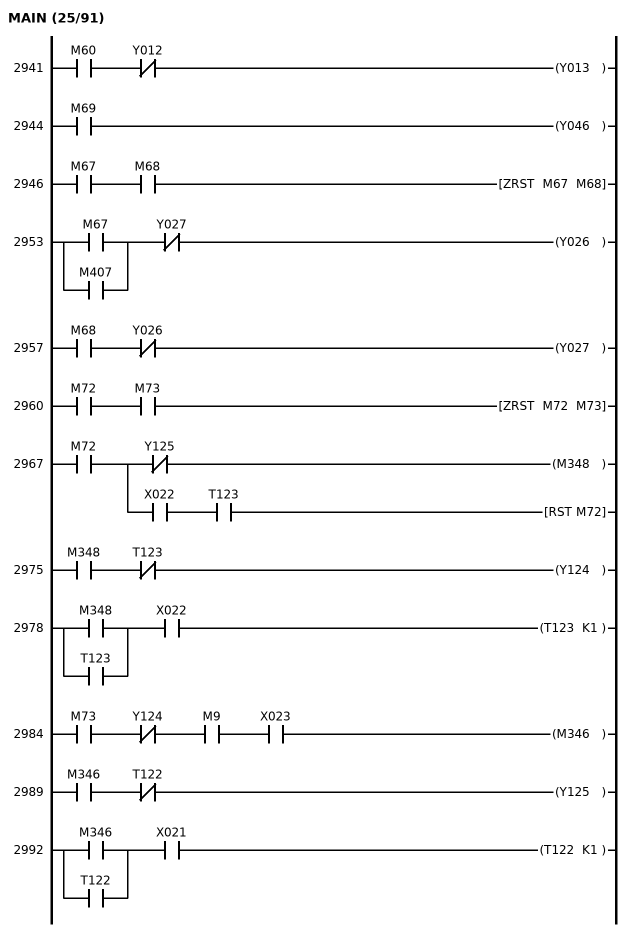
[picture p24: ladder of MAIN, rungs at steps 2941 to 2992]
2941  LD      M60
      ANI     Y012
      OUT     Y013
2944  LD      M69
      OUT     Y046
2946  LD      M67
      AND     M68
      ZRST    M67 M68
2953  LD      M67
      OR      M407
      ANI     Y027
      OUT     Y026
2957  LD      M68
      ANI     Y026
      OUT     Y027
2960  LD      M72
      AND     M73
      ZRST    M72 M73
2967  LD      M72
      MPS
      ANI     Y125
      OUT     M348
      MPP
      AND     X022
      AND     T123
      RST     M72
2975  LD      M348
      ANI     T123
      OUT     Y124
2978  LD      M348
      OR      T123
      AND     X022
      OUT     T123 K1
2984  LD      M73
      ANI     Y124
      AND     M9
      AND     X023
      OUT     M346
2989  LD      M346
      ANI     T122
      OUT     Y125
2992  LD      M346
      OR      T122
      AND     X021
      OUT     T122 K1
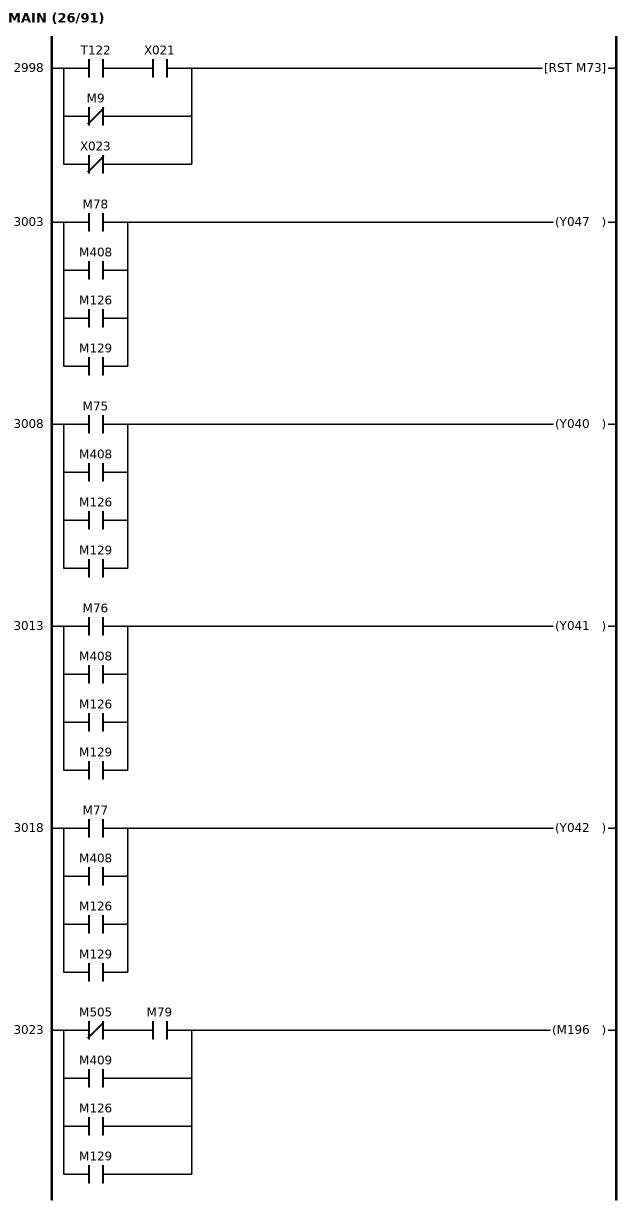
2998  LD      T122
      AND     X021
      ORI     M9
      ORI     X023
      RST     M73
3003  LD      M78
      OR      M408
      OR      M126
      OR      M129
      OUT     Y047
3008  LD      M75
      OR      M408
      OR      M126
      OR      M129
      OUT     Y040
3013  LD      M76
      OR      M408
      OR      M126
      OR      M129
      OUT     Y041
3018  LD      M77
      OR      M408
      OR      M126
      OR      M129
      OUT     Y042
3023  LDI     M505
      AND     M79
      OR      M409
      OR      M126
      OR      M129
      OUT     M196
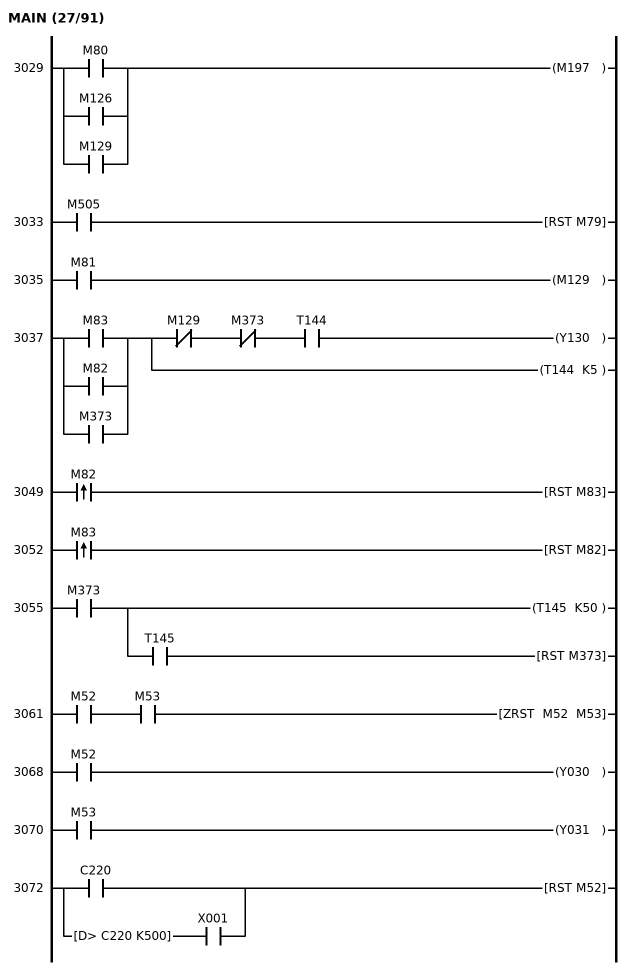
3029  LD      M80
      OR      M126
      OR      M129
      OUT     M197
3033  LD      M505
      RST     M79
3035  LD      M81
      OUT     M129
3037  LD      M83
      OR      M82
      OR      M373
      MPS
      ANI     M129
      ANI     M373
      AND     T144
      OUT     Y130
      MPP
      OUT     T144 K5
3049  LDP     M82
      RST     M83
3052  LDP     M83
      RST     M82
3055  LD      M373
      OUT     T145 K50
      AND     T145
      RST     M373
3061  LD      M52
      AND     M53
      ZRST    M52 M53
3068  LD      M52
      OUT     Y030
3070  LD      M53
      OUT     Y031
3072  LD      C220
      LDD>    C220 K500
      AND     X001
      ORB
      RST     M52
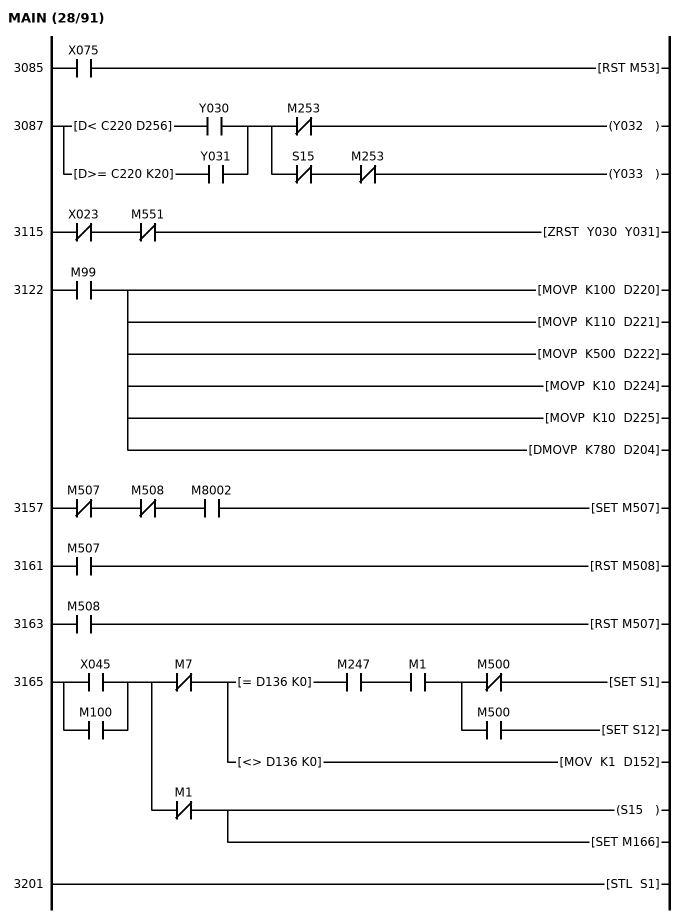
3085  LD      X075
      RST     M53
3087  LDD<    C220 D256
      AND     Y030
      LDD>=   C220 K20
      AND     Y031
      ORB
      MPS
      ANI     M253
      OUT     Y032
      MPP
      ANI     S15
      ANI     M253
      OUT     Y033
3115  LDI     X023
      ANI     M551
      ZRST    Y030 Y031
3122  LD      M99
      MOVP    K100 D220
      MOVP    K110 D221
      MOVP    K500 D222
      MOVP    K10 D224
      MOVP    K10 D225
      DMOVP   K780 D204
3157  LDI     M507
      ANI     M508
      AND     M8002
      SET     M507
3161  LD      M507
      RST     M508
3163  LD      M508
      RST     M507
3165  LD      X045
      OR      M100
      MPS
      ANI     M7
      MPS
      AND=    D136 K0
      AND     M247
      AND     M1
      MPS
      ANI     M500
      SET     S1
      MPP
      AND     M500
      SET     S12
      MPP
      AND<>   D136 K0
      MOV     K1 D152
      MPP
      ANI     M1
      OUT     S15
      SET     M166
3201  STL     S1
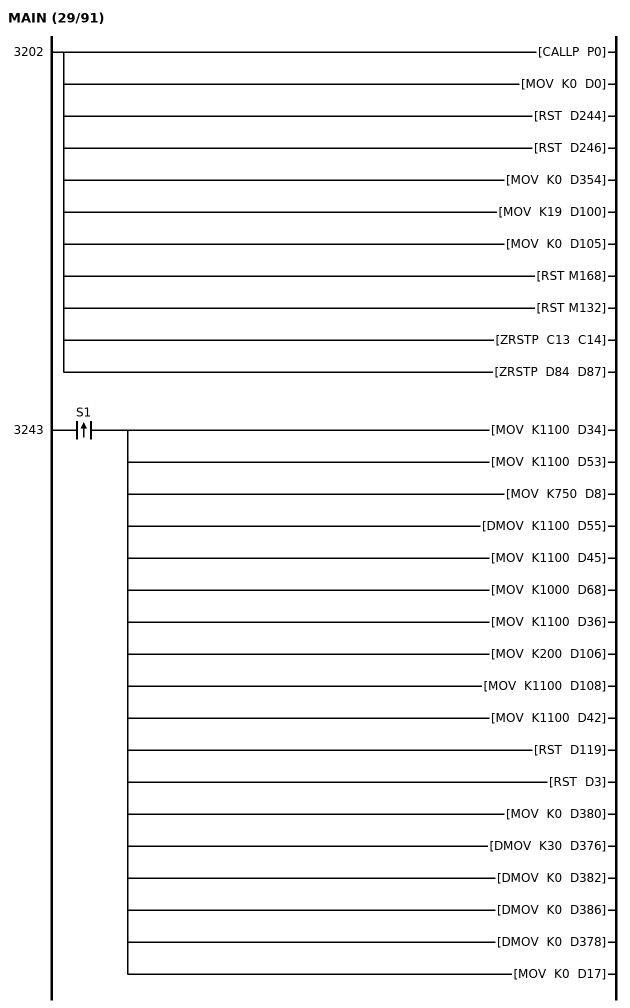
3202  CALLP   P0
      MOV     K0 D0
      RST     D244
      RST     D246
      MOV     K0 D354
      MOV     K19 D100
      MOV     K0 D105
      RST     M168
      RST     M132
      ZRSTP   C13 C14
      ZRSTP   D84 D87
3243  LDP     S1
      MOV     K1100 D34
      MOV     K1100 D53
      MOV     K750 D8
      DMOV    K1100 D55
      MOV     K1100 D45
      MOV     K1000 D68
      MOV     K1100 D36
      MOV     K200 D106
      MOV     K1100 D108
      MOV     K1100 D42
      RST     D119
      RST     D3
      MOV     K0 D380
      DMOV    K30 D376
      DMOV    K0 D382
      DMOV    K0 D386
      DMOV    K0 D378
      MOV     K0 D17
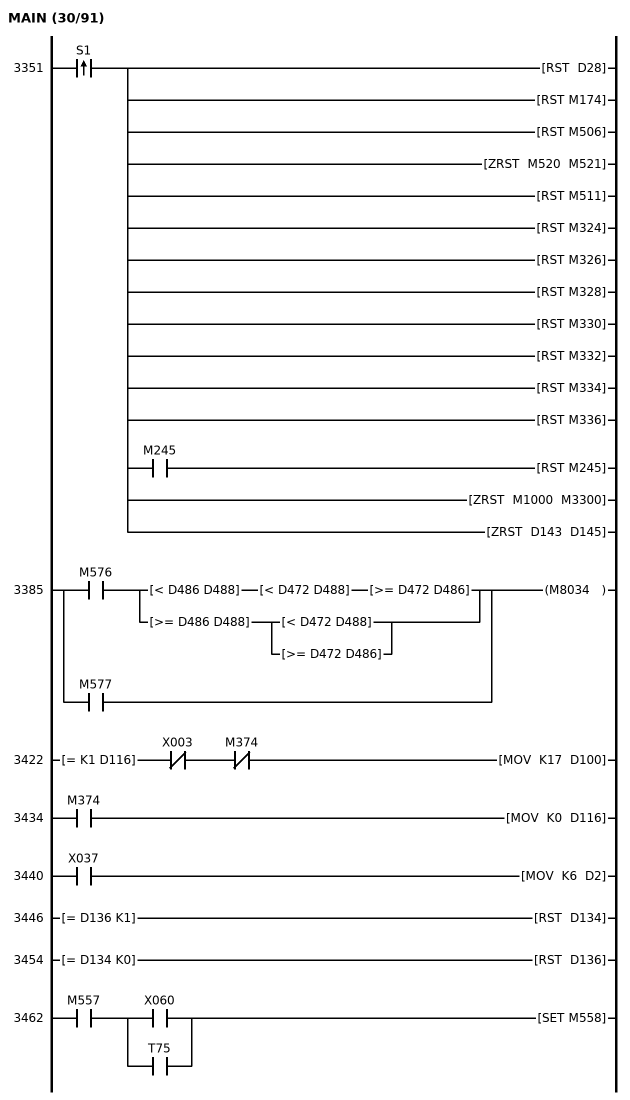
3351  LDP     S1
      RST     D28
      RST     M174
      RST     M506
      ZRST    M520 M521
      RST     M511
      RST     M324
      RST     M326
      RST     M328
      RST     M330
      RST     M332
      RST     M334
      RST     M336
      MPS
      AND     M245
      RST     M245
      MPP
      ZRST    M1000 M3300
      ZRST    D143 D145
3385  LD      M576
      LD<     D486 D488
      AND<    D472 D488
      AND>=   D472 D486
      LD>=    D486 D488
      LD<     D472 D488
      OR>=    D472 D486
      ANB
      ORB
      ANB
      OR      M577
      OUT     M8034
3422  LD=     K1 D116
      ANI     X003
      ANI     M374
      MOV     K17 D100
3434  LD      M374
      MOV     K0 D116
3440  LD      X037
      MOV     K6 D2
3446  LD=     D136 K1
      RST     D134
3454  LD=     D134 K0
      RST     D136
3462  LD      M557
      LD      X060
      OR      T75
      ANB
      SET     M558
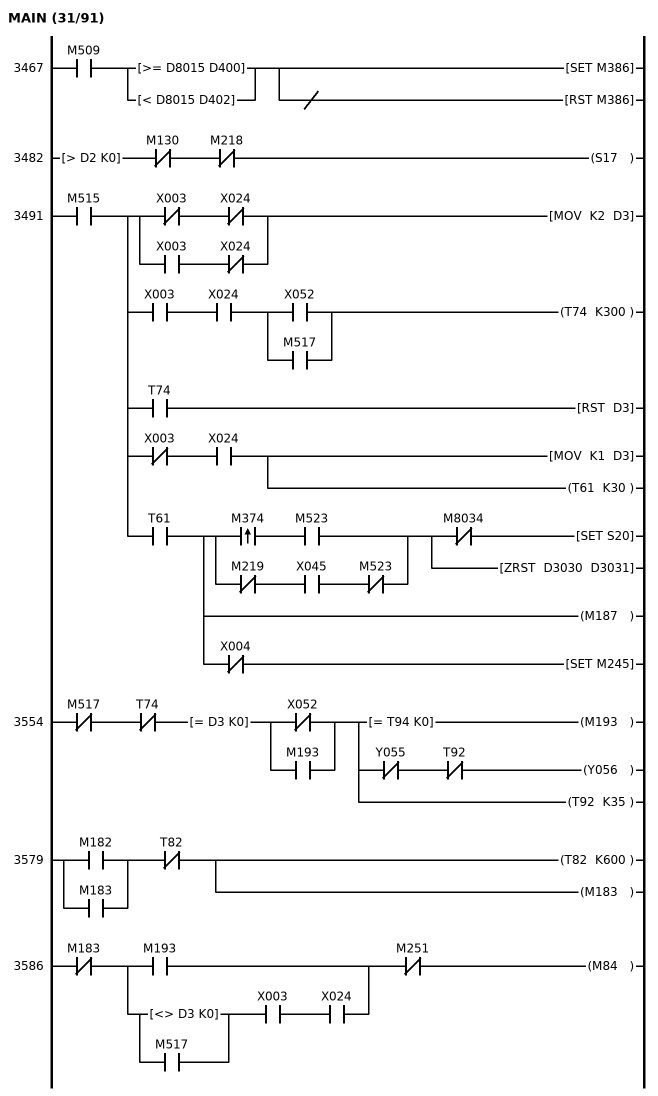
3467  LD      M509
      LD>=    D8015 D400
      OR<     D8015 D402
      ANB
      SET     M386
      INV
      RST     M386
3482  LD>     D2 K0
      ANI     M130
      ANI     M218
      OUT     S17
3491  LD      M515
      MPS
      LDI     X003
      ANI     X024
      LD      X003
      ANI     X024
      ORB
      ANB
      MOV     K2 D3
      MRD
      AND     X003
      AND     X024
      LD      X052
      OR      M517
      ANB
      OUT     T74 K300
      MRD
      AND     T74
      RST     D3
      MRD
      ANI     X003
      AND     X024
      MOV     K1 D3
      OUT     T61 K30
      MPP
      AND     T61
      MPS
      LDP     M374
      AND     M523
      LDI     M219
      AND     X045
      ANI     M523
      ORB
      ANB
      MPS
      ANI     M8034
      SET     S20
      MPP
      ZRST    D3030 D3031
      MPP
      OUT     M187
      ANI     X004
      SET     M245
3554  LDI     M517
      ANI     T74
      AND=    D3 K0
      LDI     X052
      OR      M193
      ANB
      MPS
      AND=    T94 K0
      OUT     M193
      MRD
      ANI     Y055
      ANI     T92
      OUT     Y056
      MPP
      OUT     T92 K35
3579  LD      M182
      OR      M183
      ANI     T82
      OUT     T82 K600
      OUT     M183
3586  LDI     M183
      LD      M193
      LD<>    D3 K0
      OR      M517
      AND     X003
      AND     X024
      ORB
      ANB
      ANI     M251
      OUT     M84
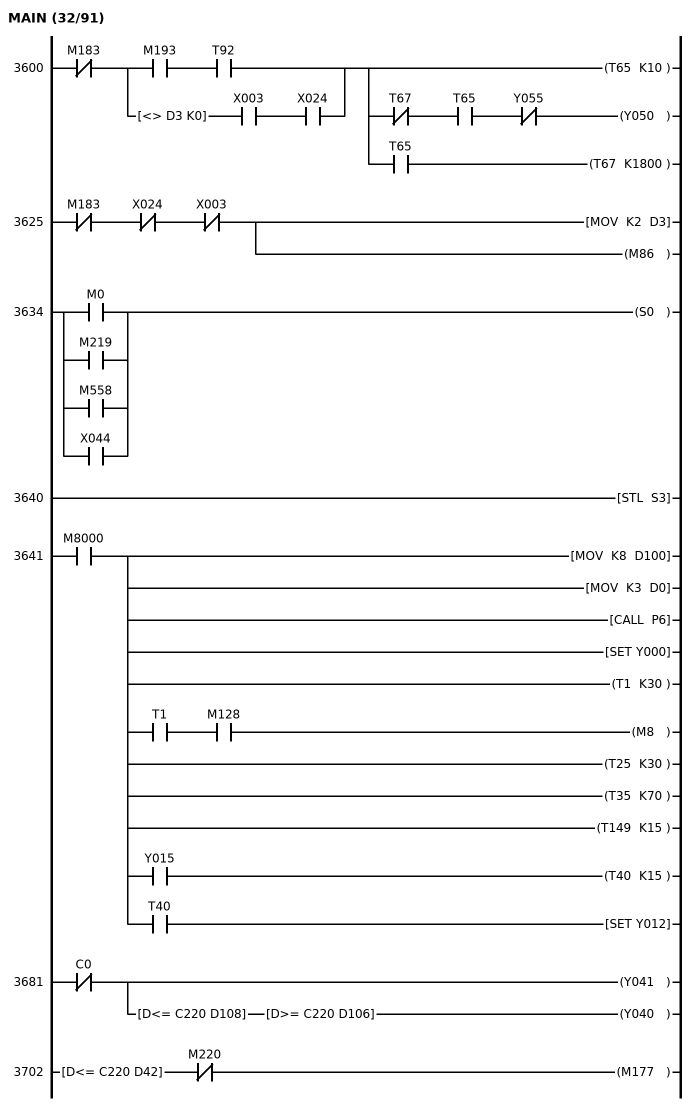
3600  LDI     M183
      LD      M193
      AND     T92
      LD<>    D3 K0
      AND     X003
      AND     X024
      ORB
      ANB
      OUT     T65 K10
      MPS
      ANI     T67
      AND     T65
      ANI     Y055
      OUT     Y050
      MPP
      AND     T65
      OUT     T67 K1800
3625  LDI     M183
      ANI     X024
      ANI     X003
      MOV     K2 D3
      OUT     M86
3634  LD      M0
      OR      M219
      OR      M558
      OR      X044
      OUT     S0
3640  STL     S3
3641  LD      M8000
      MOV     K8 D100
      MOV     K3 D0
      CALL    P6
      SET     Y000
      OUT     T1 K30
      MPS
      AND     T1
      AND     M128
      OUT     M8
      MPP
      OUT     T25 K30
      OUT     T35 K70
      OUT     T149 K15
      MPS
      AND     Y015
      OUT     T40 K15
      MPP
      AND     T40
      SET     Y012
3681  LDI     C0
      OUT     Y041
      ANDD<=  C220 D108
      ANDD>=  C220 D106
      OUT     Y040
3702  LDD<=   C220 D42
      ANI     M220
      OUT     M177
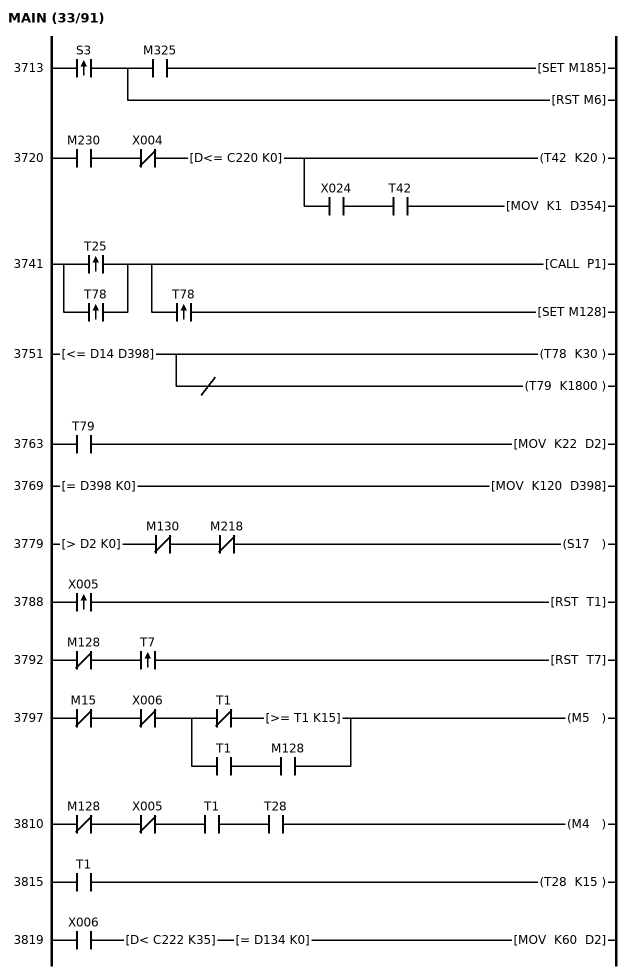
3713  LDP     S3
      MPS
      AND     M325
      SET     M185
      MPP
      RST     M6
3720  LD      M230
      ANI     X004
      ANDD<=  C220 K0
      OUT     T42 K20
      AND     X024
      AND     T42
      MOV     K1 D354
3741  LDP     T25
      ORP     T78
      CALL    P1
      ANDP    T78
      SET     M128
3751  LD<=    D14 D398
      OUT     T78 K30
      INV
      OUT     T79 K1800
3763  LD      T79
      MOV     K22 D2
3769  LD=     D398 K0
      MOV     K120 D398
3779  LD>     D2 K0
      ANI     M130
      ANI     M218
      OUT     S17
3788  LDP     X005
      RST     T1
3792  LDI     M128
      ANDP    T7
      RST     T7
3797  LDI     M15
      ANI     X006
      LDI     T1
      AND>=   T1 K15
      LD      T1
      AND     M128
      ORB
      ANB
      OUT     M5
3810  LDI     M128
      ANI     X005
      AND     T1
      AND     T28
      OUT     M4
3815  LD      T1
      OUT     T28 K15
3819  LD      X006
      ANDD<   C222 K35
      AND=    D134 K0
      MOV     K60 D2
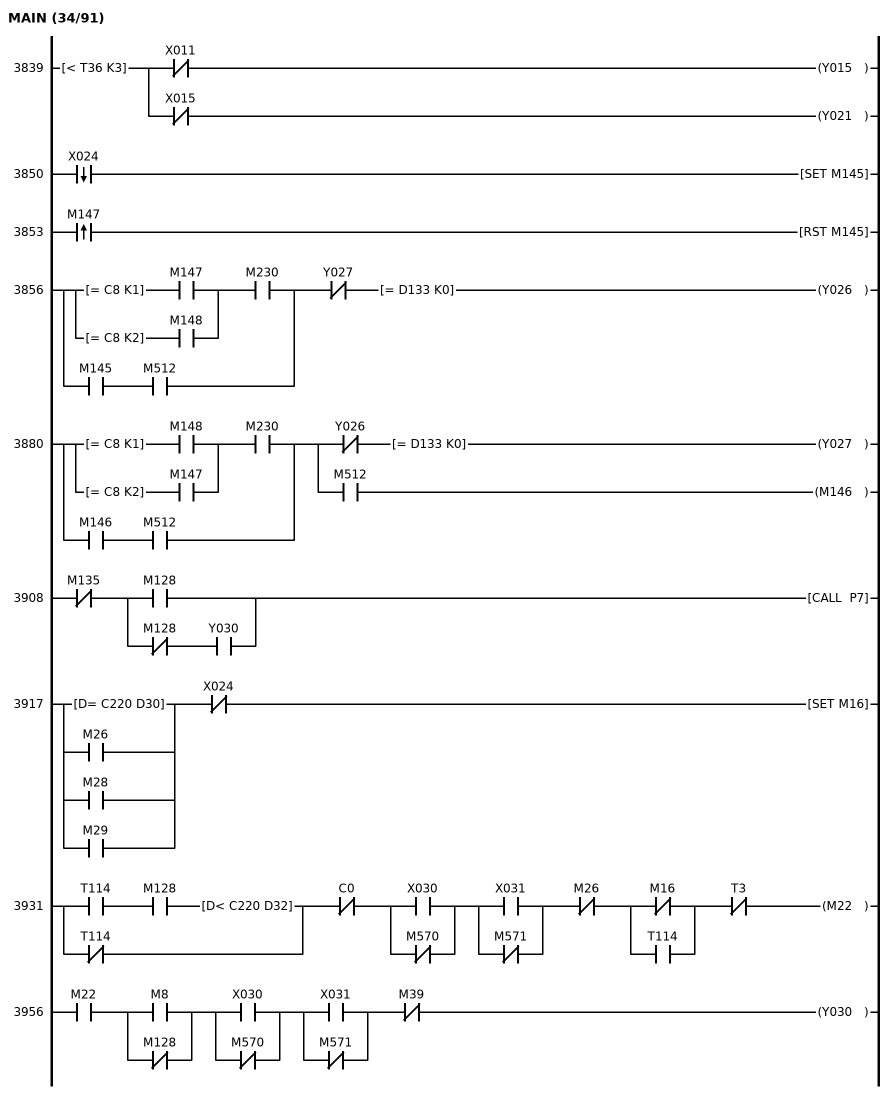
3839  LD<     T36 K3
      MPS
      ANI     X011
      OUT     Y015
      MPP
      ANI     X015
      OUT     Y021
3850  LDF     X024
      SET     M145
3853  LDP     M147
      RST     M145
3856  LD=     C8 K1
      AND     M147
      LD=     C8 K2
      AND     M148
      ORB
      AND     M230
      LD      M145
      AND     M512
      ORB
      ANI     Y027
      AND=    D133 K0
      OUT     Y026
3880  LD=     C8 K1
      AND     M148
      LD=     C8 K2
      AND     M147
      ORB
      AND     M230
      LD      M146
      AND     M512
      ORB
      MPS
      ANI     Y026
      AND=    D133 K0
      OUT     Y027
      MPP
      AND     M512
      OUT     M146
3908  LDI     M135
      LD      M128
      LDI     M128
      AND     Y030
      ORB
      ANB
      CALL    P7
3917  LDD=    C220 D30
      OR      M26
      OR      M28
      OR      M29
      ANI     X024
      SET     M16
3931  LD      T114
      AND     M128
      ANDD<   C220 D32
      ORI     T114
      ANI     C0
      LD      X030
      ORI     M570
      ANB
      LD      X031
      ORI     M571
      ANB
      ANI     M26
      LDI     M16
      OR      T114
      ANB
      ANI     T3
      OUT     M22
3956  LD      M22
      LD      M8
      ORI     M128
      ANB
      LD      X030
      ORI     M570
      ANB
      LD      X031
      ORI     M571
      ANB
      ANI     M39
      OUT     Y030
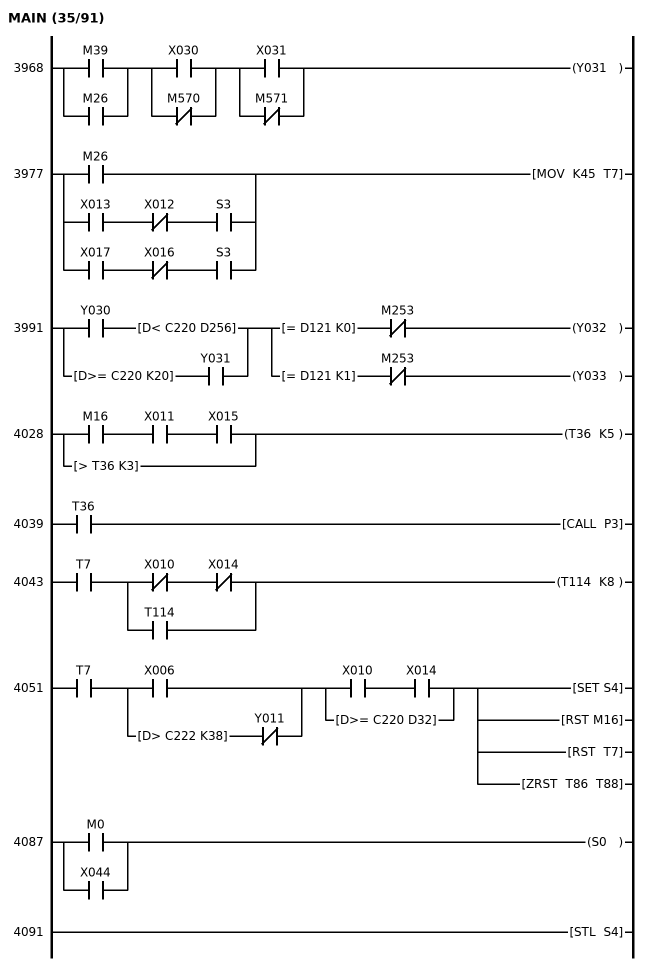
3968  LD      M39
      OR      M26
      LD      X030
      ORI     M570
      ANB
      LD      X031
      ORI     M571
      ANB
      OUT     Y031
3977  LD      M26
      LD      X013
      ANI     X012
      AND     S3
      ORB
      LD      X017
      ANI     X016
      AND     S3
      ORB
      MOV     K45 T7
3991  LD      Y030
      ANDD<   C220 D256
      LDD>=   C220 K20
      AND     Y031
      ORB
      MPS
      AND=    D121 K0
      ANI     M253
      OUT     Y032
      MPP
      AND=    D121 K1
      ANI     M253
      OUT     Y033
4028  LD      M16
      AND     X011
      AND     X015
      OR>     T36 K3
      OUT     T36 K5
4039  LD      T36
      CALL    P3
4043  LD      T7
      LDI     X010
      ANI     X014
      OR      T114
      ANB
      OUT     T114 K8
4051  LD      T7
      LD      X006
      LDD>    C222 K38
      ANI     Y011
      ORB
      ANB
      LD      X010
      AND     X014
      ORD>=   C220 D32
      ANB
      SET     S4
      RST     M16
      RST     T7
      ZRST    T86 T88
4087  LD      M0
      OR      X044
      OUT     S0
4091  STL     S4
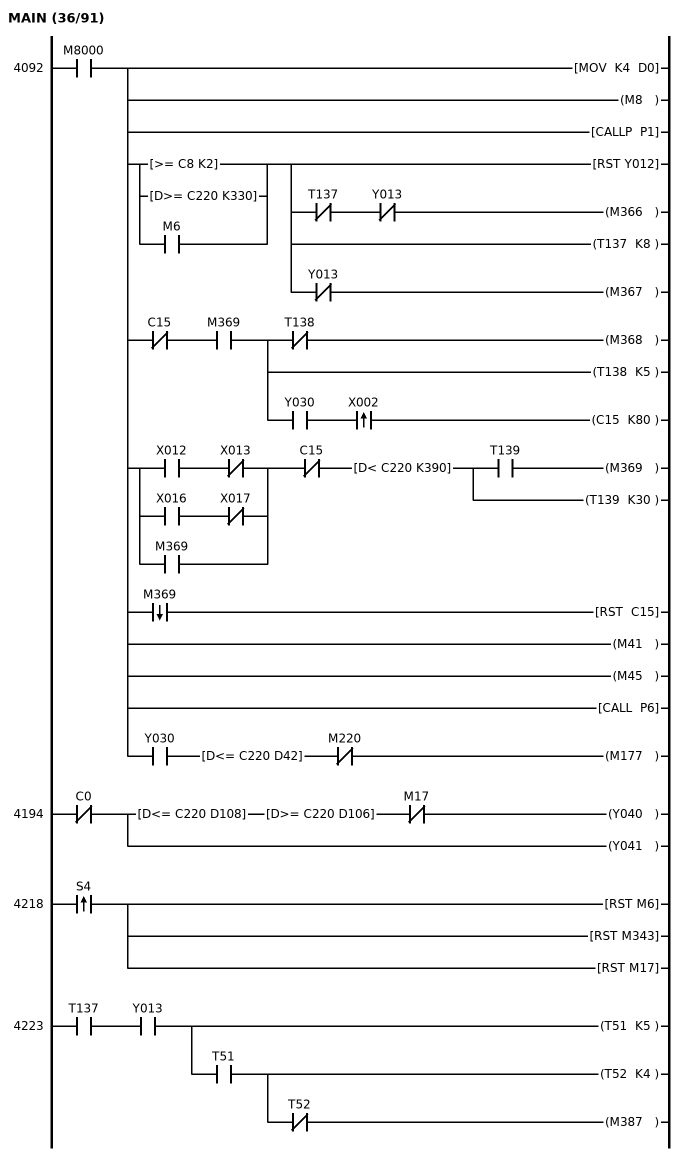
4092  LD      M8000
      MOV     K4 D0
      OUT     M8
      CALLP   P1
      MPS
      LD>=    C8 K2
      ORD>=   C220 K330
      OR      M6
      ANB
      RST     Y012
      MPS
      ANI     T137
      ANI     Y013
      OUT     M366
      MPP
      OUT     T137 K8
      ANI     Y013
      OUT     M367
      MRD
      ANI     C15
      AND     M369
      MPS
      ANI     T138
      OUT     M368
      MPP
      OUT     T138 K5
      AND     Y030
      ANDP    X002
      OUT     C15 K80
      MRD
      LD      X012
      ANI     X013
      LD      X016
      ANI     X017
      ORB
      OR      M369
      ANB
      ANI     C15
      ANDD<   C220 K390
      MPS
      AND     T139
      OUT     M369
      MPP
      OUT     T139 K30
      MRD
      ANDF    M369
      RST     C15
      MPP
      OUT     M41
      OUT     M45
      CALL    P6
      AND     Y030
      ANDD<=  C220 D42
      ANI     M220
      OUT     M177
4194  LDI     C0
      MPS
      ANDD<=  C220 D108
      ANDD>=  C220 D106
      ANI     M17
      OUT     Y040
      MPP
      OUT     Y041
4218  LDP     S4
      RST     M6
      RST     M343
      RST     M17
4223  LD      T137
      AND     Y013
      OUT     T51 K5
      AND     T51
      OUT     T52 K4
      ANI     T52
      OUT     M387
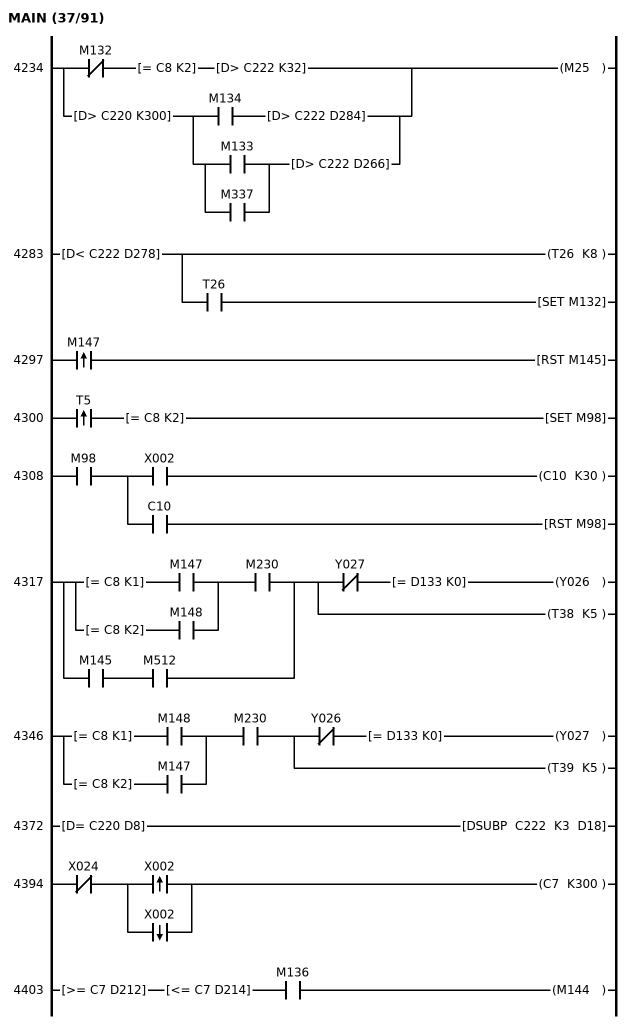
4234  LDI     M132
      AND=    C8 K2
      ANDD>   C222 K32
      LDD>    C220 K300
      LD      M134
      ANDD>   C222 D284
      LD      M133
      OR      M337
      ANDD>   C222 D266
      ORB
      ANB
      ORB
      OUT     M25
4283  LDD<    C222 D278
      OUT     T26 K8
      AND     T26
      SET     M132
4297  LDP     M147
      RST     M145
4300  LDP     T5
      AND=    C8 K2
      SET     M98
4308  LD      M98
      MPS
      AND     X002
      OUT     C10 K30
      MPP
      AND     C10
      RST     M98
4317  LD=     C8 K1
      AND     M147
      LD=     C8 K2
      AND     M148
      ORB
      AND     M230
      LD      M145
      AND     M512
      ORB
      MPS
      ANI     Y027
      AND=    D133 K0
      OUT     Y026
      MPP
      OUT     T38 K5
4346  LD=     C8 K1
      AND     M148
      LD=     C8 K2
      AND     M147
      ORB
      AND     M230
      MPS
      ANI     Y026
      AND=    D133 K0
      OUT     Y027
      MPP
      OUT     T39 K5
4372  LDD=    C220 D8
      DSUBP   C222 K3 D18
4394  LDI     X024
      LDP     X002
      ORF     X002
      ANB
      OUT     C7 K300
4403  LD>=    C7 D212
      AND<=   C7 D214
      AND     M136
      OUT     M144
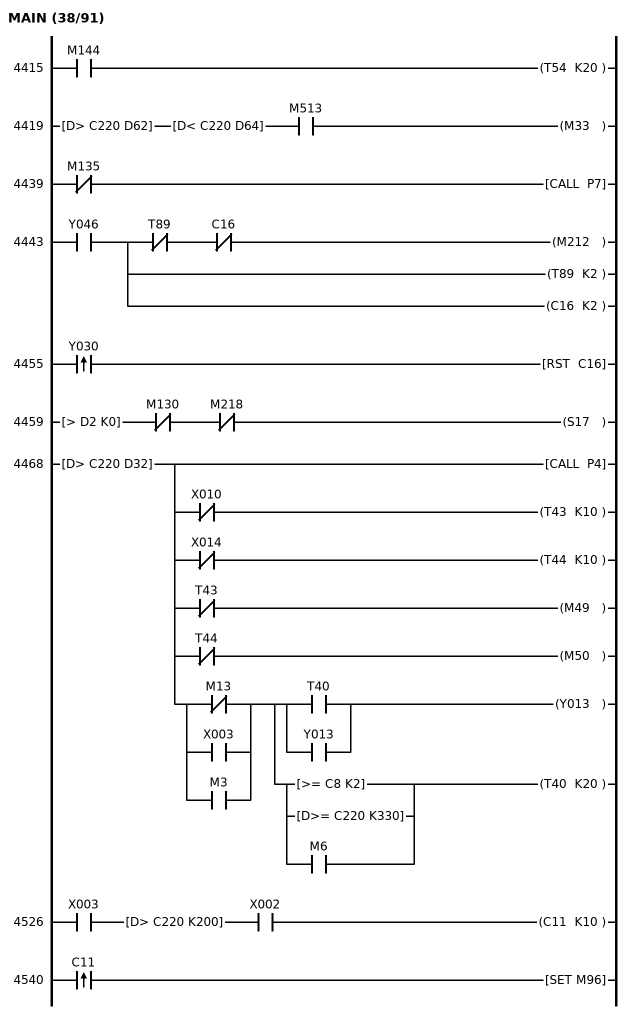
4415  LD      M144
      OUT     T54 K20
4419  LDD>    C220 D62
      ANDD<   C220 D64
      AND     M513
      OUT     M33
4439  LDI     M135
      CALL    P7
4443  LD      Y046
      MPS
      ANI     T89
      ANI     C16
      OUT     M212
      MPP
      OUT     T89 K2
      OUT     C16 K2
4455  LDP     Y030
      RST     C16
4459  LD>     D2 K0
      ANI     M130
      ANI     M218
      OUT     S17
4468  LDD>    C220 D32
      CALL    P4
      MPS
      ANI     X010
      OUT     T43 K10
      MRD
      ANI     X014
      OUT     T44 K10
      MRD
      ANI     T43
      OUT     M49
      MRD
      ANI     T44
      OUT     M50
      MPP
      LDI     M13
      OR      X003
      OR      M3
      ANB
      MPS
      LD      T40
      OR      Y013
      ANB
      OUT     Y013
      MPP
      LD>=    C8 K2
      ORD>=   C220 K330
      OR      M6
      ANB
      OUT     T40 K20
4526  LD      X003
      ANDD>   C220 K200
      AND     X002
      OUT     C11 K10
4540  LDP     C11
      SET     M96
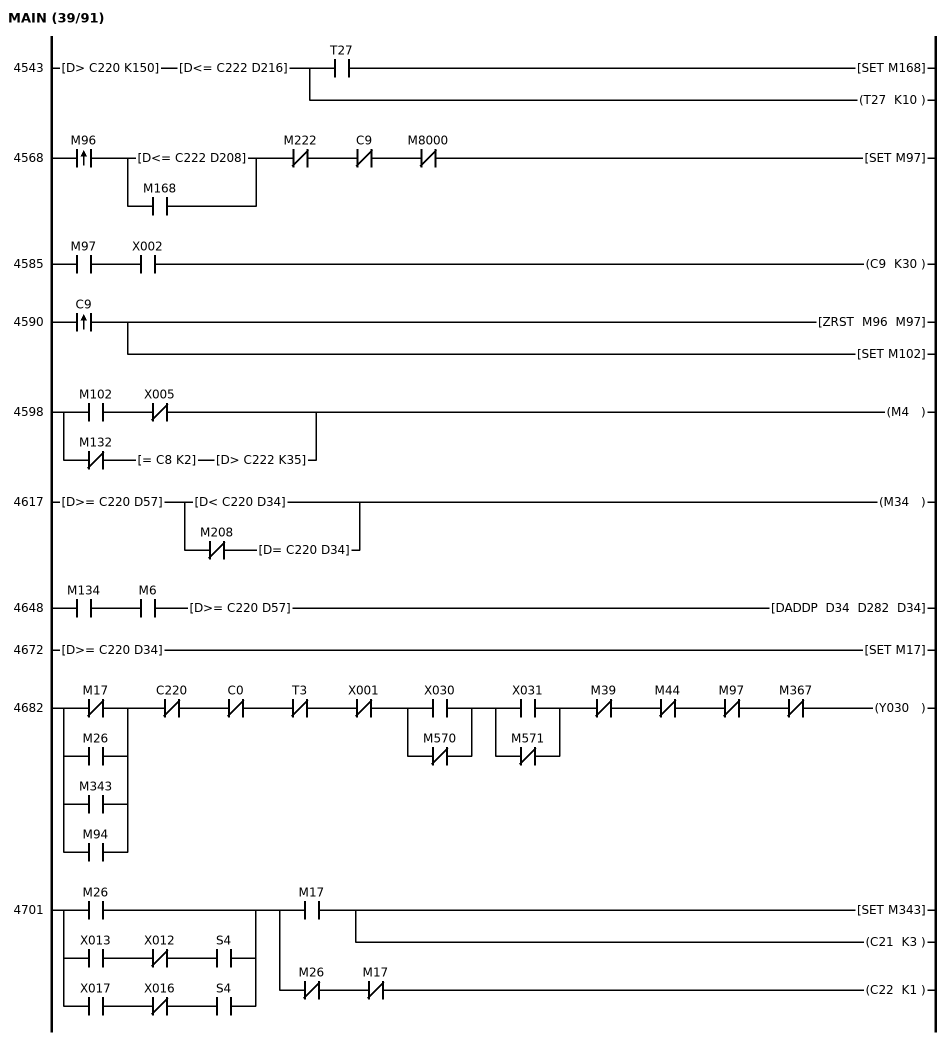
4543  LDD>    C220 K150
      ANDD<=  C222 D216
      MPS
      AND     T27
      SET     M168
      MPP
      OUT     T27 K10
4568  LDP     M96
      LDD<=   C222 D208
      OR      M168
      ANB
      ANI     M222
      ANI     C9
      ANI     M8000
      SET     M97
4585  LD      M97
      AND     X002
      OUT     C9 K30
4590  LDP     C9
      ZRST    M96 M97
      SET     M102
4598  LD      M102
      ANI     X005
      LDI     M132
      AND=    C8 K2
      ANDD>   C222 K35
      ORB
      OUT     M4
4617  LDD>=   C220 D57
      LDD<    C220 D34
      LDI     M208
      ANDD=   C220 D34
      ORB
      ANB
      OUT     M34
4648  LD      M134
      AND     M6
      ANDD>=  C220 D57
      DADDP   D34 D282 D34
4672  LDD>=   C220 D34
      SET     M17
4682  LDI     M17
      OR      M26
      OR      M343
      OR      M94
      ANI     C220
      ANI     C0
      ANI     T3
      ANI     X001
      LD      X030
      ORI     M570
      ANB
      LD      X031
      ORI     M571
      ANB
      ANI     M39
      ANI     M44
      ANI     M97
      ANI     M367
      OUT     Y030
4701  LD      M26
      LD      X013
      ANI     X012
      AND     S4
      ORB
      LD      X017
      ANI     X016
      AND     S4
      ORB
      MPS
      AND     M17
      SET     M343
      OUT     C21 K3
      MPP
      ANI     M26
      ANI     M17
      OUT     C22 K1
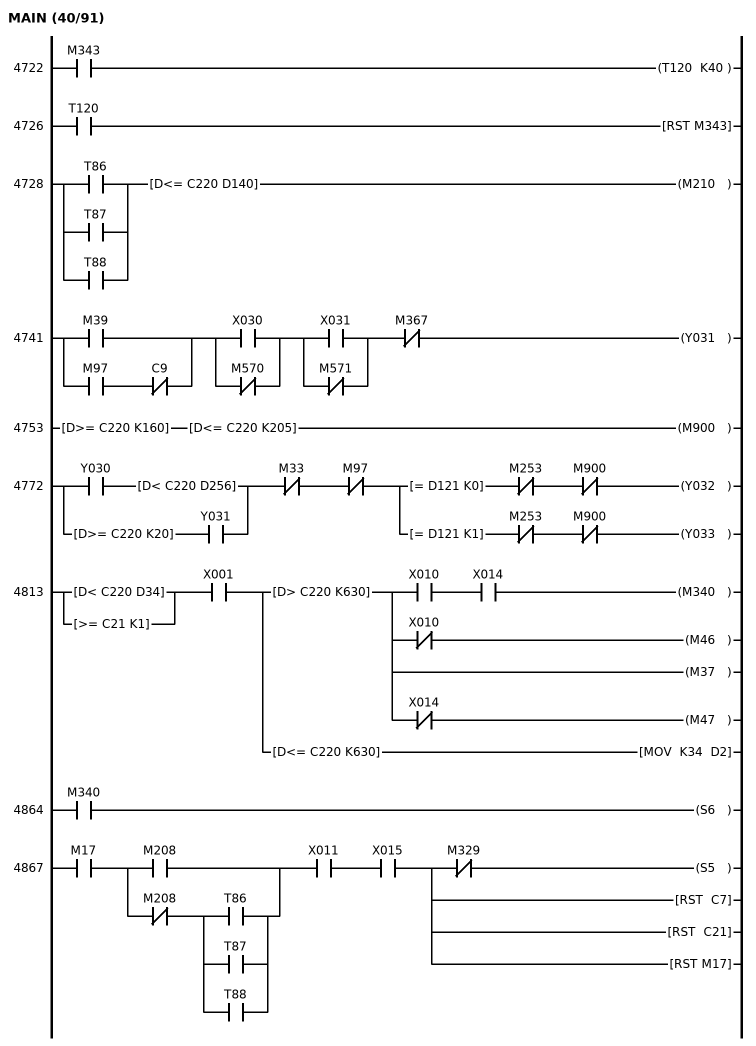
4722  LD      M343
      OUT     T120 K40
4726  LD      T120
      RST     M343
4728  LD      T86
      OR      T87
      OR      T88
      ANDD<=  C220 D140
      OUT     M210
4741  LD      M39
      LD      M97
      ANI     C9
      ORB
      LD      X030
      ORI     M570
      ANB
      LD      X031
      ORI     M571
      ANB
      ANI     M367
      OUT     Y031
4753  LDD>=   C220 K160
      ANDD<=  C220 K205
      OUT     M900
4772  LD      Y030
      ANDD<   C220 D256
      LDD>=   C220 K20
      AND     Y031
      ORB
      ANI     M33
      ANI     M97
      MPS
      AND=    D121 K0
      ANI     M253
      ANI     M900
      OUT     Y032
      MPP
      AND=    D121 K1
      ANI     M253
      ANI     M900
      OUT     Y033
4813  LDD<    C220 D34
      OR>=    C21 K1
      AND     X001
      MPS
      ANDD>   C220 K630
      MPS
      AND     X010
      AND     X014
      OUT     M340
      MRD
      ANI     X010
      OUT     M46
      MPP
      OUT     M37
      ANI     X014
      OUT     M47
      MPP
      ANDD<=  C220 K630
      MOV     K34 D2
4864  LD      M340
      OUT     S6
4867  LD      M17
      LD      M208
      LDI     M208
      LD      T86
      OR      T87
      OR      T88
      ANB
      ORB
      ANB
      AND     X011
      AND     X015
      MPS
      ANI     M329
      OUT     S5
      MPP
      RST     C7
      RST     C21
      RST     M17
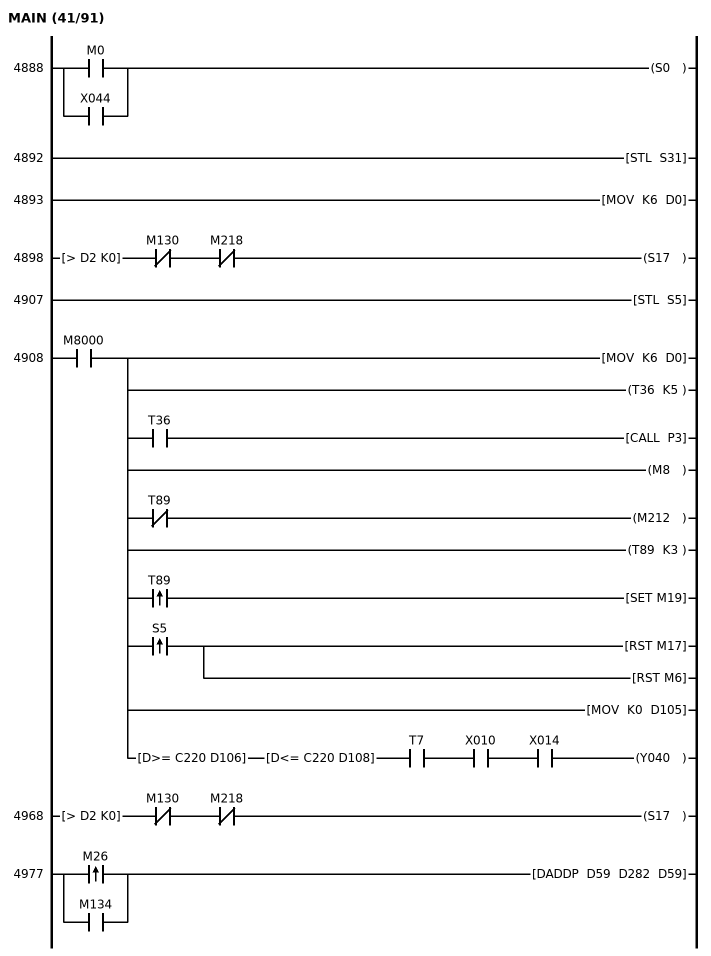
4888  LD      M0
      OR      X044
      OUT     S0
4892  STL     S31
4893  MOV     K6 D0
4898  LD>     D2 K0
      ANI     M130
      ANI     M218
      OUT     S17
4907  STL     S5
4908  LD      M8000
      MOV     K6 D0
      OUT     T36 K5
      MPS
      AND     T36
      CALL    P3
      MPP
      OUT     M8
      MPS
      ANI     T89
      OUT     M212
      MPP
      OUT     T89 K3
      MPS
      ANDP    T89
      SET     M19
      MRD
      ANDP    S5
      RST     M17
      RST     M6
      MPP
      MOV     K0 D105
      ANDD>=  C220 D106
      ANDD<=  C220 D108
      AND     T7
      AND     X010
      AND     X014
      OUT     Y040
4968  LD>     D2 K0
      ANI     M130
      ANI     M218
      OUT     S17
4977  LDP     M26
      OR      M134
      DADDP   D59 D282 D59
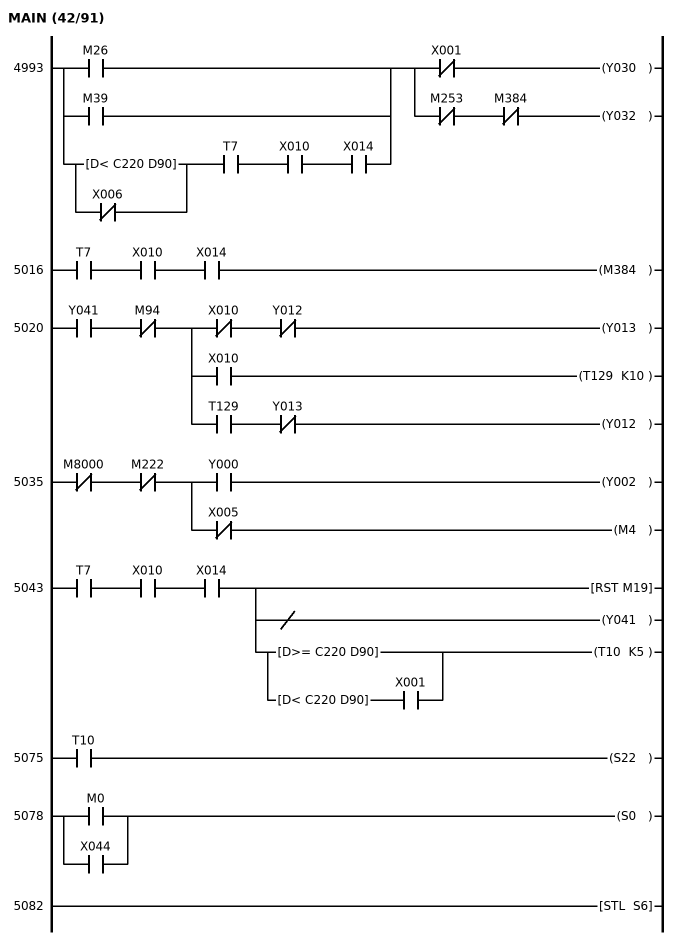
4993  LD      M26
      OR      M39
      LDD<    C220 D90
      ORI     X006
      AND     T7
      AND     X010
      AND     X014
      ORB
      MPS
      ANI     X001
      OUT     Y030
      MPP
      ANI     M253
      ANI     M384
      OUT     Y032
5016  LD      T7
      AND     X010
      AND     X014
      OUT     M384
5020  LD      Y041
      ANI     M94
      MPS
      ANI     X010
      ANI     Y012
      OUT     Y013
      MRD
      AND     X010
      OUT     T129 K10
      MPP
      AND     T129
      ANI     Y013
      OUT     Y012
5035  LDI     M8000
      ANI     M222
      MPS
      AND     Y000
      OUT     Y002
      MPP
      ANI     X005
      OUT     M4
5043  LD      T7
      AND     X010
      AND     X014
      RST     M19
      MPS
      INV
      OUT     Y041
      MPP
      LDD>=   C220 D90
      LDD<    C220 D90
      AND     X001
      ORB
      ANB
      OUT     T10 K5
5075  LD      T10
      OUT     S22
5078  LD      M0
      OR      X044
      OUT     S0
5082  STL     S6
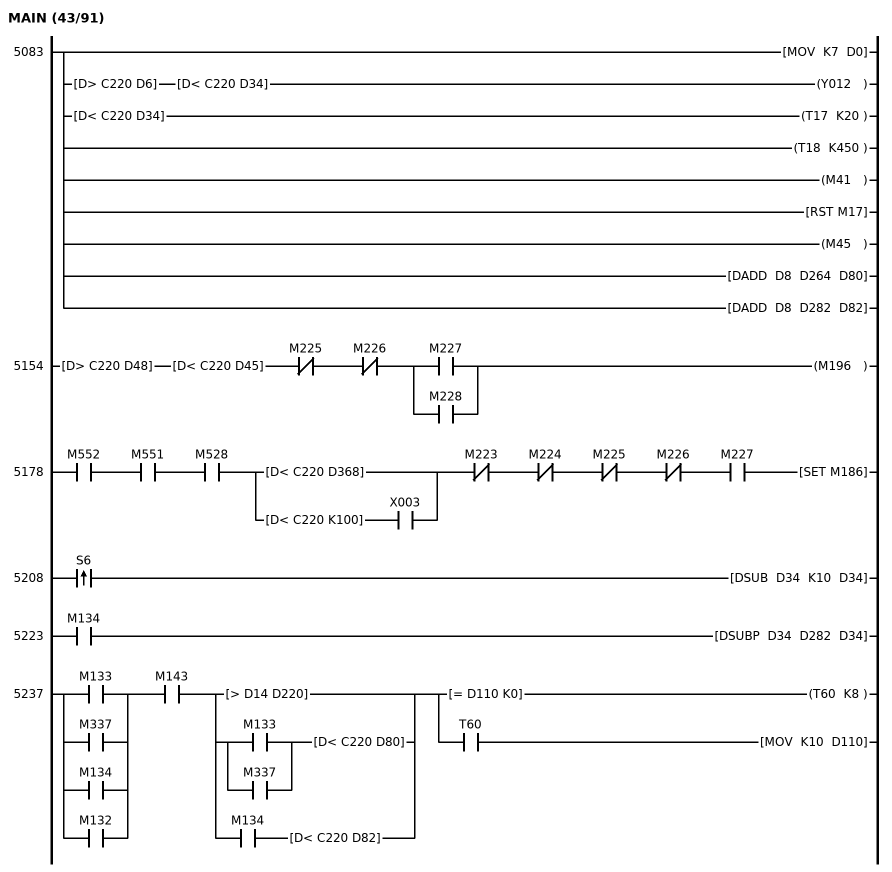
5083  MOV     K7 D0
      MPS
      ANDD>   C220 D6
      ANDD<   C220 D34
      OUT     Y012
      MRD
      ANDD<   C220 D34
      OUT     T17 K20
      MPP
      OUT     T18 K450
      OUT     M41
      RST     M17
      OUT     M45
      DADD    D8 D264 D80
      DADD    D8 D282 D82
5154  LDD>    C220 D48
      ANDD<   C220 D45
      ANI     M225
      ANI     M226
      LD      M227
      OR      M228
      ANB
      OUT     M196
5178  LD      M552
      AND     M551
      AND     M528
      LDD<    C220 D368
      LDD<    C220 K100
      AND     X003
      ORB
      ANB
      ANI     M223
      ANI     M224
      ANI     M225
      ANI     M226
      AND     M227
      SET     M186
5208  LDP     S6
      DSUB    D34 K10 D34
5223  LD      M134
      DSUBP   D34 D282 D34
5237  LD      M133
      OR      M337
      OR      M134
      OR      M132
      AND     M143
      LD>     D14 D220
      LD      M133
      OR      M337
      ANDD<   C220 D80
      ORB
      LD      M134
      ANDD<   C220 D82
      ORB
      ANB
      MPS
      AND=    D110 K0
      OUT     T60 K8
      MPP
      AND     T60
      MOV     K10 D110
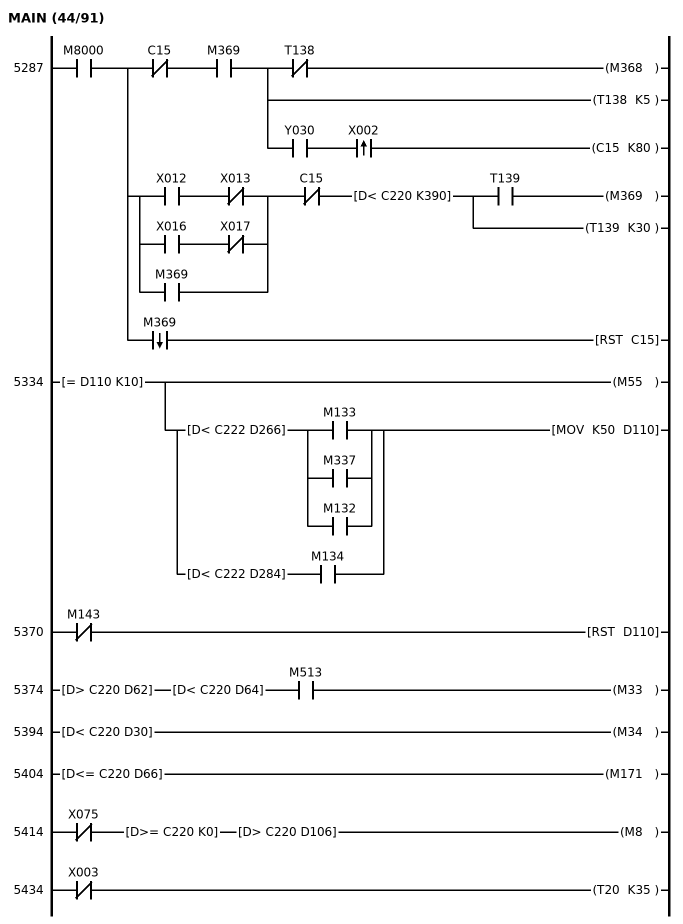
5287  LD      M8000
      MPS
      ANI     C15
      AND     M369
      MPS
      ANI     T138
      OUT     M368
      MPP
      OUT     T138 K5
      AND     Y030
      ANDP    X002
      OUT     C15 K80
      MRD
      LD      X012
      ANI     X013
      LD      X016
      ANI     X017
      ORB
      OR      M369
      ANB
      ANI     C15
      ANDD<   C220 K390
      MPS
      AND     T139
      OUT     M369
      MPP
      OUT     T139 K30
      MPP
      ANDF    M369
      RST     C15
5334  LD=     D110 K10
      OUT     M55
      LDD<    C222 D266
      LD      M133
      OR      M337
      OR      M132
      ANB
      LDD<    C222 D284
      AND     M134
      ORB
      ANB
      MOV     K50 D110
5370  LDI     M143
      RST     D110
5374  LDD>    C220 D62
      ANDD<   C220 D64
      AND     M513
      OUT     M33
5394  LDD<    C220 D30
      OUT     M34
5404  LDD<=   C220 D66
      OUT     M171
5414  LDI     X075
      ANDD>=  C220 K0
      ANDD>   C220 D106
      OUT     M8
5434  LDI     X003
      OUT     T20 K35
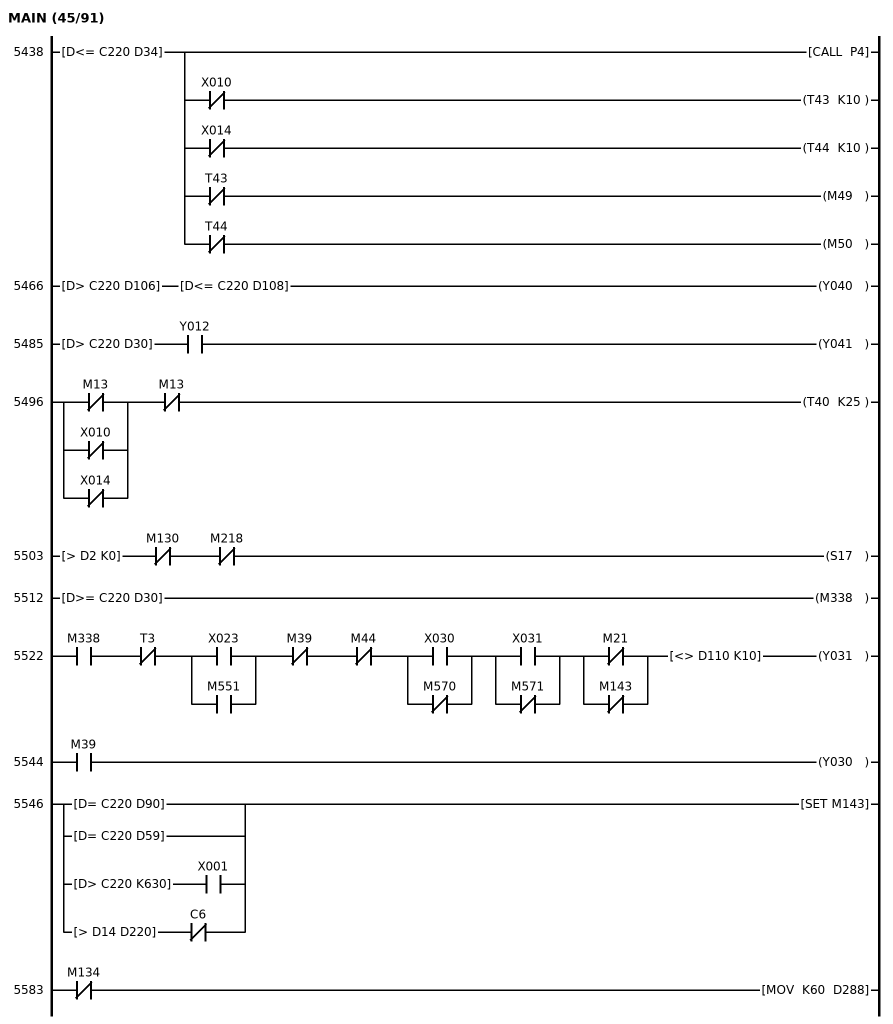
5438  LDD<=   C220 D34
      CALL    P4
      MPS
      ANI     X010
      OUT     T43 K10
      MRD
      ANI     X014
      OUT     T44 K10
      MRD
      ANI     T43
      OUT     M49
      MPP
      ANI     T44
      OUT     M50
5466  LDD>    C220 D106
      ANDD<=  C220 D108
      OUT     Y040
5485  LDD>    C220 D30
      AND     Y012
      OUT     Y041
5496  LDI     M13
      ORI     X010
      ORI     X014
      ANI     M13
      OUT     T40 K25
5503  LD>     D2 K0
      ANI     M130
      ANI     M218
      OUT     S17
5512  LDD>=   C220 D30
      OUT     M338
5522  LD      M338
      ANI     T3
      LD      X023
      OR      M551
      ANB
      ANI     M39
      ANI     M44
      LD      X030
      ORI     M570
      ANB
      LD      X031
      ORI     M571
      ANB
      LDI     M21
      ORI     M143
      ANB
      AND<>   D110 K10
      OUT     Y031
5544  LD      M39
      OUT     Y030
5546  LDD=    C220 D90
      ORD=    C220 D59
      LDD>    C220 K630
      AND     X001
      ORB
      LD>     D14 D220
      ANI     C6
      ORB
      SET     M143
5583  LDI     M134
      MOV     K60 D288
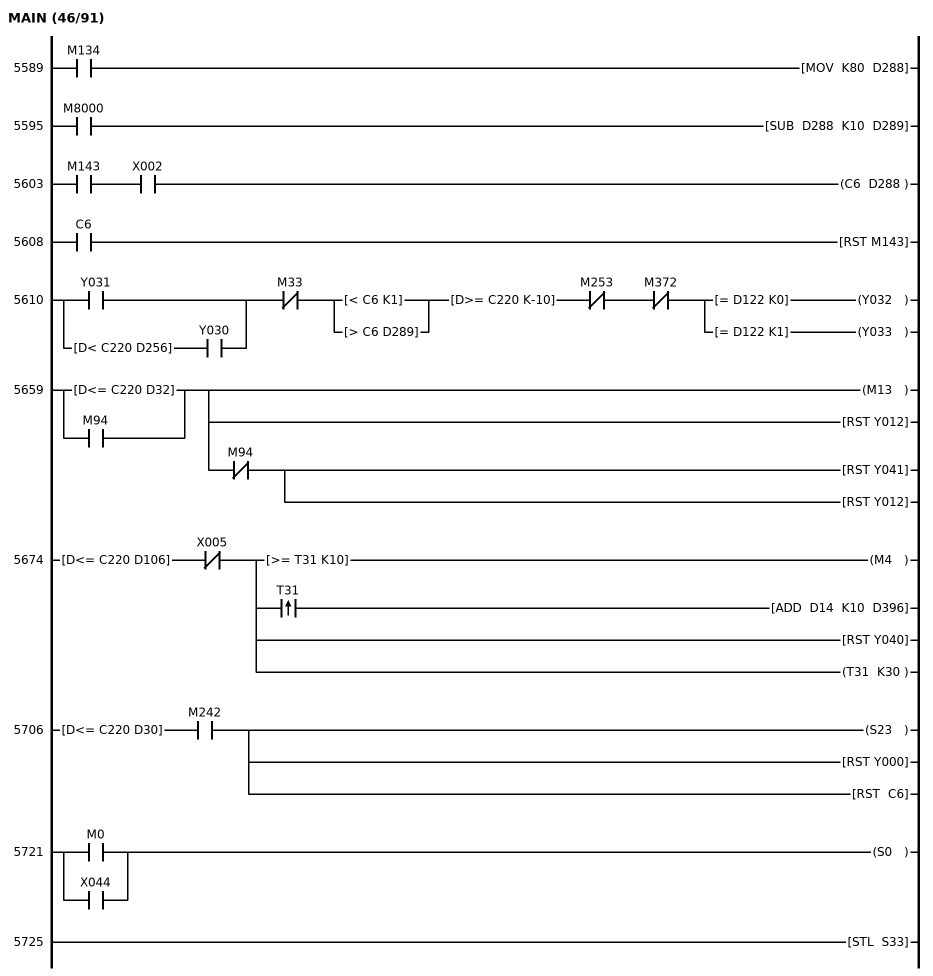
5589  LD      M134
      MOV     K80 D288
5595  LD      M8000
      SUB     D288 K10 D289
5603  LD      M143
      AND     X002
      OUT     C6 D288
5608  LD      C6
      RST     M143
5610  LD      Y031
      LDD<    C220 D256
      AND     Y030
      ORB
      ANI     M33
      LD<     C6 K1
      OR>     C6 D289
      ANB
      ANDD>=  C220 K-10
      ANI     M253
      ANI     M372
      MPS
      AND=    D122 K0
      OUT     Y032
      MPP
      AND=    D122 K1
      OUT     Y033
5659  LDD<=   C220 D32
      OR      M94
      OUT     M13
      RST     Y012
      ANI     M94
      RST     Y041
      RST     Y012
5674  LDD<=   C220 D106
      ANI     X005
      MPS
      AND>=   T31 K10
      OUT     M4
      MRD
      ANDP    T31
      ADD     D14 K10 D396
      MPP
      RST     Y040
      OUT     T31 K30
5706  LDD<=   C220 D30
      AND     M242
      OUT     S23
      RST     Y000
      RST     C6
5721  LD      M0
      OR      X044
      OUT     S0
5725  STL     S33
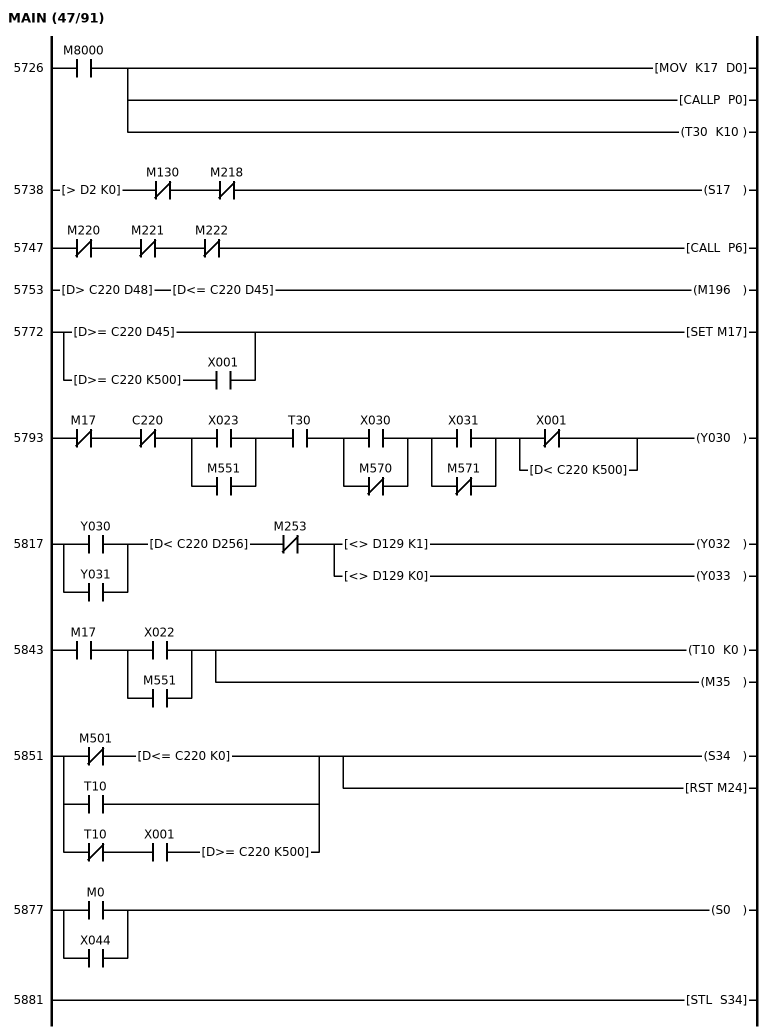
5726  LD      M8000
      MOV     K17 D0
      CALLP   P0
      OUT     T30 K10
5738  LD>     D2 K0
      ANI     M130
      ANI     M218
      OUT     S17
5747  LDI     M220
      ANI     M221
      ANI     M222
      CALL    P6
5753  LDD>    C220 D48
      ANDD<=  C220 D45
      OUT     M196
5772  LDD>=   C220 D45
      LDD>=   C220 K500
      AND     X001
      ORB
      SET     M17
5793  LDI     M17
      ANI     C220
      LD      X023
      OR      M551
      ANB
      AND     T30
      LD      X030
      ORI     M570
      ANB
      LD      X031
      ORI     M571
      ANB
      LDI     X001
      ORD<    C220 K500
      ANB
      OUT     Y030
5817  LD      Y030
      OR      Y031
      ANDD<   C220 D256
      ANI     M253
      MPS
      AND<>   D129 K1
      OUT     Y032
      MPP
      AND<>   D129 K0
      OUT     Y033
5843  LD      M17
      LD      X022
      OR      M551
      ANB
      OUT     T10 K0
      OUT     M35
5851  LDI     M501
      ANDD<=  C220 K0
      OR      T10
      LDI     T10
      AND     X001
      ANDD>=  C220 K500
      ORB
      OUT     S34
      RST     M24
5877  LD      M0
      OR      X044
      OUT     S0
5881  STL     S34
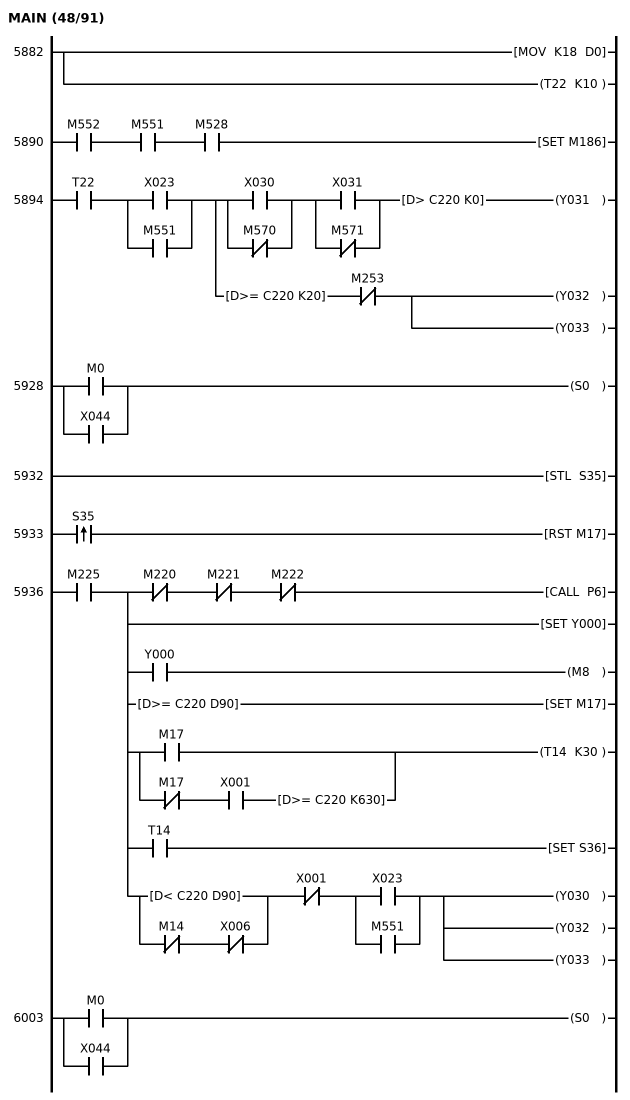
5882  MOV     K18 D0
      OUT     T22 K10
5890  LD      M552
      AND     M551
      AND     M528
      SET     M186
5894  LD      T22
      LD      X023
      OR      M551
      ANB
      MPS
      LD      X030
      ORI     M570
      ANB
      LD      X031
      ORI     M571
      ANB
      ANDD>   C220 K0
      OUT     Y031
      MPP
      ANDD>=  C220 K20
      ANI     M253
      OUT     Y032
      OUT     Y033
5928  LD      M0
      OR      X044
      OUT     S0
5932  STL     S35
5933  LDP     S35
      RST     M17
5936  LD      M225
      MPS
      ANI     M220
      ANI     M221
      ANI     M222
      CALL    P6
      MPP
      SET     Y000
      MPS
      AND     Y000
      OUT     M8
      MRD
      ANDD>=  C220 D90
      SET     M17
      MRD
      LD      M17
      LDI     M17
      AND     X001
      ANDD>=  C220 K630
      ORB
      ANB
      OUT     T14 K30
      MRD
      AND     T14
      SET     S36
      MPP
      LDD<    C220 D90
      LDI     M14
      ANI     X006
      ORB
      ANB
      ANI     X001
      LD      X023
      OR      M551
      ANB
      OUT     Y030
      OUT     Y032
      OUT     Y033
6003  LD      M0
      OR      X044
      OUT     S0
